Fanuc KAREL source: kb00014.KL

-- PROVISIONAL review KL for V1013-1; original PC SHA256 807387370bf03192a888e2aece3824ccbce43a92425736c26e7b74a460263e7f
-- Incomplete behavior may be omitted. Consult companion uncertainty JSON. Do not deploy.
PROGRAM KB00014
%NOLOCKGROUP
BEGIN
  -- UNRESOLVED_PC offsets 5-21; opcodes 27,22,31,23
  -- UNRESOLVED_PC offsets 26-30; opcodes 7F
END KB00014
